Fanuc KAREL source: compact_preamble.KL

PROGRAM KA00001
%NOLOCKGROUP
VAR
SRC:INTEGER;DST:INTEGER
BEGIN
SRC=2
DST=SRC
END KA00001
